FUNCTION_BLOCK FB_Equipment
VAR_INPUT
END_VAR
VAR_OUTPUT
END_VAR
VAR
END_VAR

END_FUNCTION_BLOCK

(* stored: Version 1.1.0.1
   POU FB_Equipment: Id {f1dba864-9346-4d69-9b08-e58db36c0188}, SpecialFunc None *)
